Fanuc KAREL source: kt00339.KL

-- PROVISIONAL review KL for V940-1; original PC SHA256 9a0a5599f54b1b1ea19fd1132495f1be4cca87a5c5dbb7e1c39fc89be9432569
-- Incomplete behavior may be omitted. Consult companion uncertainty JSON. Do not deploy.
PROGRAM KT00339
%NOLOCKGROUP
VAR
  I2 : INTEGER
  OUT : BOOLEAN
-- UNRESOLVED_DECL Y1 type=002018
BEGIN
  -- V9_ZERO_TABLE_METADATA_HINT layout=0001; no indexed target words; source/name/runtime held
  -- UNRESOLVED_PC offsets 5-19; opcodes 2E,22,9D,33,B2
  -- UNRESOLVED_PC offsets 24-35; opcodes 2E,23
  -- UNRESOLVED_PC offsets 40-62; opcodes 22,9D,33,B1,21,59,23
  -- UNRESOLVED_PC offsets 67-71; opcodes 7F
END KT00339
